(* Schneider Machine Expert - Basic project modbus_07_write_read_mw_fc23_il_only, file version 3.0.0.0 *)
(* ProjectInformations: Name=New project *)

HARDWARE
  Cpu 0: TM200CE40T
  EthernetConfiguration: NetworkName=M200, IpAllocationMode=FixedAddress, IpAddress=0.0.0.0, SubnetMask=0.0.0.0
  SerialLineConfiguration: Baud=Baud19200, Parity=ParityEven, DataBits=DataBits8, StopBits=StopBits1, PhysicalMedium=PhysicalMediumRs485, TransmissionMode=TransmissionModeModbusRtu, SlaveId=1, Addressing=MasterAddressing
  MastTask: UsePeriodScanMode=false, PeriodScan=100
  FastTask: Period=255
  CpuBehavior: StartingMode=StartAsPreviousState, AutoSaveRamOnEeprom=true, WatchdogPeriod=250

SYMBOLS  (address, symbol, comment, settings)
  %WRITE_READ_VAR0   [Link(Value(FBComLinkParameterEnums=SerialLine1)), RemoteDeviceId(Value(int=1)), Timeout(Value(int=100)), ObjType(Value(FBComObjTypeParameterEnums=MW)), FirstWriteObj(Value(int=17)), WriteQuantity(Value(int=2)), IndexDataOut(Value(int=300)), FirstReadObj(Value(int=41)), ReadQuantity(Value(int=3)), IndexDataIn(Value(int=400))]

POU Generated C++ - EXPERIMENTAL
  (* SectionNumber=0 *)

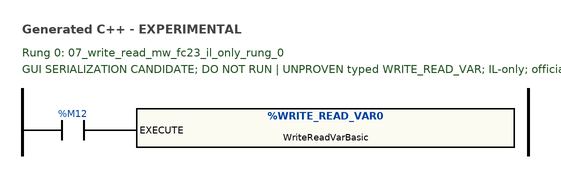

// Rung 0: 07_write_read_mw_fc23_il_only_rung_0
// GUI SERIALIZATION CANDIDATE; DO NOT RUN | UNPROVEN typed WRITE_READ_VAR; IL-only; official Ladder conversion required
  BLK %WRITE_READ_VAR0
  LD %M12
  EXECUTE
  END_BLK
  // as ST:
  //   %WRITE_READ_VAR0(EXECUTE := %M12);
